Omron CX-Programmer project NewProject (CX-Programmer 9.73)

# PLC UAS_AUTOCLAVE: CJ2M CPU31
I/O table (CPU CJ2M-CPU31): rack 0 slot 0 CJ1W-AD041-V1; rack 0 slot 1 CJ1W-DA041; rack 0 slot 2 CJ1W-TC001; rack 0 slot 3 CJ1W-ID211; rack 0 slot 4 CJ1W-OC211; rack 0 slot 11 CJ2M-EIP21

## Global symbols (name address type ; comment)
0.00 BOOL  ; START
0.01 BOOL  ; STOP
100.01 BOOL  ; DANGER
100.02 BOOL  ; SUHU BOILER
100.03 BOOL  ; TEKANAN BOILER
100.05 BOOL  ; BOILER ON/OFF
100.06 BOOL  ; SUHU AUTOCLAVE
100.07 BOOL  ; TEKANAN AUTOCLAVE
100.08 BOOL  ; STERILIZING
100.09 BOOL  ; RELEASE
100.10 BOOL  ; COOLING
100.11 BOOL  ; SAFE
100.12 BOOL  ; CONNECT
1.01 BOOL  ; DANGER
1.02 BOOL  ; SUHU BOILER
1.03 BOOL  ; TEKANAN BOILER
1.05 BOOL  ; BOILER ON/OFF (HEATING)
1.06 BOOL  ; SUHU AUTOCLAVE
1.07 BOOL  ; TEKANAN AUTOCLAVE
1.08 BOOL  ; STERILIZING
1.09 BOOL  ; RELEASE
1.10 BOOL  ; COOLING
1.11 BOOL  ; SAFE
1.12 BOOL  ; CONNECT
D0 CHANNEL  ; SUHU BOILER
D1 CHANNEL  ; TEKANAN BOILER
D2 CHANNEL  ; SUHU AUTOCLAVE
D3 CHANNEL  ; SET POINT SUHU AUTOCLAVE
D4 CHANNEL  ; TEKANAN AUTOCLAVE
D5 CHANNEL  ; SET POINT TEKANAN AUTOCLAVE
D6 CHANNEL  ; TIMER STERILIZING
D7 CHANNEL  ; TIMER RELEASE
D8 CHANNEL  ; TIMER COOLING
T0 CHANNEL  ; TIMER STERILIZING
T0000 BOOL  ; TIMER STERILIZING
T0001 BOOL  ; TIMER RELEASE
T0002 BOOL  ; TIMER COOLING
T1 CHANNEL  ; TIMER RELEASE
T2 CHANNEL  ; TIMER COOLING

## Program NewProgram1 (cyclic task 0)

### Section Section1

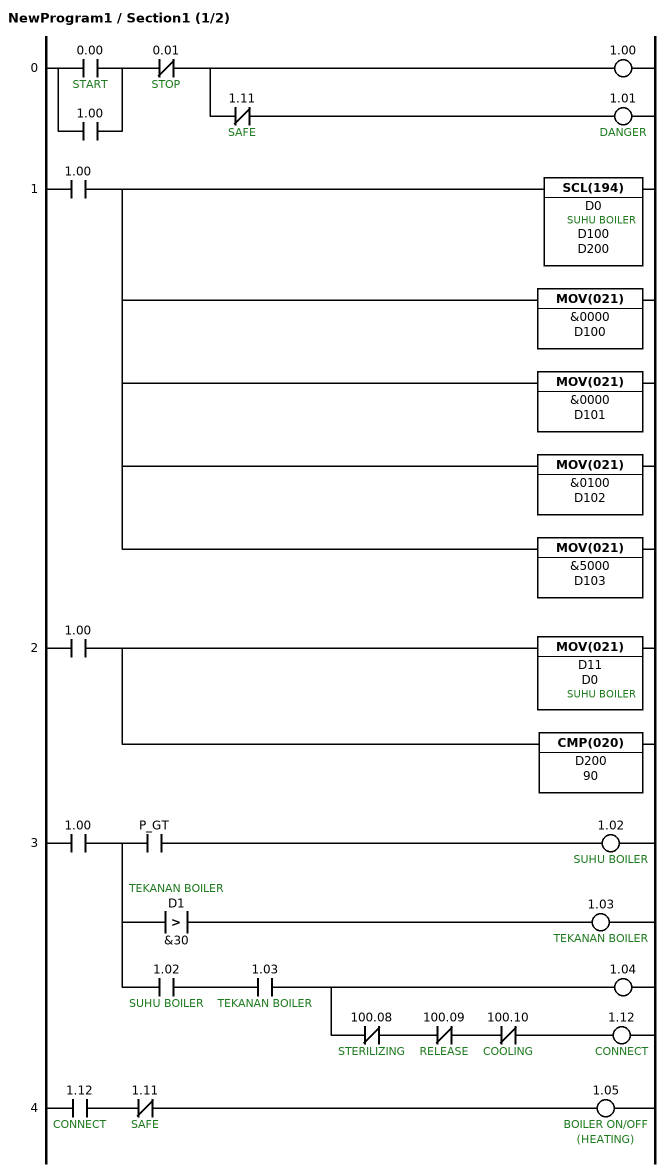
; rung 0
LD 0.00  ; START
OR 1.00
ANDNOT 0.01  ; STOP
OUT 1.00
ANDNOT 1.11  ; SAFE
OUT 1.01  ; DANGER
; rung 1
LD 1.00
SCL(194) D0 D100 D200  ; SUHU BOILER
MOV(021) &0000 D100
MOV(021) &0000 D101
MOV(021) &0100 D102
MOV(021) &5000 D103
; rung 2
LD 1.00
MOV(021) D11 D0  ; SUHU BOILER
CMP(020) D200 90
; rung 3
LD 1.00
OUT TR0
AND P_GT
OUT 1.02  ; SUHU BOILER
LD TR0
AND>(320) D1 &30  ; TEKANAN BOILER
OUT 1.03  ; TEKANAN BOILER
LD TR0
AND 1.02  ; SUHU BOILER
AND 1.03  ; TEKANAN BOILER
OUT 1.04
ANDNOT 100.08  ; STERILIZING
ANDNOT 100.09  ; RELEASE
ANDNOT 100.10  ; COOLING
OUT 1.12  ; CONNECT
; rung 4
LD 1.12  ; CONNECT
ANDNOT 1.11  ; SAFE
OUT 1.05  ; BOILER ON/OFF (HEATING)

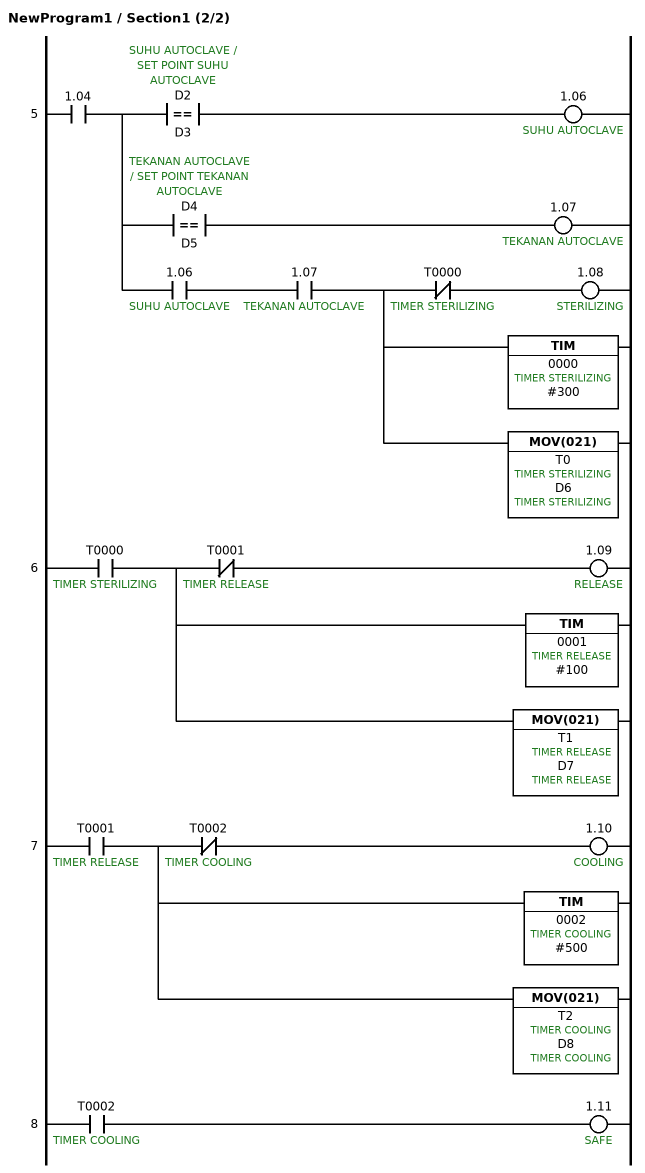
; rung 5
LD 1.04
OUT TR0
AND=(300) D2 D3  ; SUHU AUTOCLAVE, SET POINT SUHU AUTOCLAVE
OUT 1.06  ; SUHU AUTOCLAVE
LD TR0
AND=(300) D4 D5  ; TEKANAN AUTOCLAVE, SET POINT TEKANAN AUTOCLAVE
OUT 1.07  ; TEKANAN AUTOCLAVE
LD TR0
AND 1.06  ; SUHU AUTOCLAVE
AND 1.07  ; TEKANAN AUTOCLAVE
OUT TR0
ANDNOT T0000  ; TIMER STERILIZING
OUT 1.08  ; STERILIZING
LD TR0
TIM 0000 #300  ; TIMER STERILIZING
MOV(021) T0 D6  ; TIMER STERILIZING
; rung 6
LD T0000  ; TIMER STERILIZING
OUT TR0
ANDNOT T0001  ; TIMER RELEASE
OUT 1.09  ; RELEASE
LD TR0
TIM 0001 #100  ; TIMER RELEASE
MOV(021) T1 D7  ; TIMER RELEASE
; rung 7
LD T0001  ; TIMER RELEASE
OUT TR0
ANDNOT T0002  ; TIMER COOLING
OUT 1.10  ; COOLING
LD TR0
TIM 0002 #500  ; TIMER COOLING
MOV(021) T2 D8  ; TIMER COOLING
; rung 8
LD T0002  ; TIMER COOLING
OUT 1.11  ; SAFE

### Section END
; rung 0
END(001)